(* IEC 61131-3 sources: trust-platform/examples/twincat-ads/src, 2 files *)

(* ---- config.st ---- *)
CONFIGURATION Config
RESOURCE MainRes ON PLC
    TASK MainTask (INTERVAL := T#10ms, PRIORITY := 1);
    PROGRAM Main WITH MainTask : Main;
END_RESOURCE
END_CONFIGURATION

(* ---- Main.st ---- *)
PROGRAM Main
VAR
    heartbeat : DINT;
END_VAR
    heartbeat := heartbeat + 1;
END_PROGRAM
